# EPICS substitutions: db/Beckhoff_7XXX/ecmcEP7211-0034_OPT_touchProbe.substitutions
file "ecmcEL72XX_TP.template"
{
  pattern {CH_ID}
          {01   }
}
